{region 'Documentation'}
(*!
<summary>Checks that at least one selected bit is TRUE.</summary>
*)
{endregion}
FUNCTION_BLOCK AssertContainsTrue_Word EXTENDS AssertionBase
VAR_INPUT
    IN : WORD; //! Actual bitfield.
    Mask : WORD := 16#FFFF; //! Selects evaluated bits; defaults to all bits. An empty mask produces Error during evaluation.
END_VAR

SUPER^();

{region 'Documentation'}
(*!
<summary>Rejects an empty mask before checking for a matching selected bit.</summary>
*)
{endregion}
METHOD PROTECTED Assert
VAR
    Message : STRING(GVL_Constants.MessageLength);
    MaskText : STRING(GVL_Constants.AssertionValueLength);
    ActualText : STRING(GVL_Constants.AssertionValueLength);
END_VAR
VAR CONSTANT
    NoMask : WORD := 16#00;
    HexDigitCount : USINT := 4;
END_VAR
IF NOT EvaluationActive THEN
    RETURN;
END_IF;

IF Result = E_Result.Error THEN
    RETURN;
END_IF;

IF Mask = NoMask THEN
    MaskText := CreateAssertionTextValue_Hex(Value := WORD_TO_LWORD(Mask),
        DigitCount := HexDigitCount);
    Message := CONCAT('Assertion error: mask must not be empty. Mask = ',
        MaskText);
    Message := CONCAT(Message, '.');
    Error(Message := Message);
    RETURN;
END_IF;

IF Result = E_Result.Failed THEN
    RETURN;
END_IF;

IF (IN AND Mask) = NoMask THEN
    MaskText := CreateAssertionTextValue_Hex(Value := WORD_TO_LWORD(Mask),
        DigitCount := HexDigitCount);
    ActualText := CreateAssertionTextValue_Hex(Value := WORD_TO_LWORD(IN),
        DigitCount := HexDigitCount);
    Message := CONCAT('Assertion failed: no selected bit is TRUE. Mask = ',
        MaskText);
    Message := CONCAT(Message, ', Actual = ');
    Message := CONCAT(Message, ActualText);
    Message := CONCAT(Message, '.');
    Fail(Message := Message);
    RETURN;
END_IF;

Pass();
END_METHOD

END_FUNCTION_BLOCK

(* stored: Version 1.1.0.1
   POU AssertContainsTrue_Word: Id {d3f53912-88fa-4635-bfe6-0a4b6b28a83c}, SpecialFunc None
   Folder Internal: Id {54567756-ca7f-45c6-bd0e-212520f07541}
   Method Assert: Id {531fd97a-1a57-465d-8f47-0e66a90b4f17} *)
